// TIA Portal V21 export
// export: Created 2026-11-10T19:11:41.20904Z, ExportSetting WithDefaults, DisplayName Totally Integrated Automation Portal, DisplayVersion V21 Update 3, DisplayName STEP 7 Professional, DisplayVersion V21 Update 3, DisplayName STEP 7 Safety, DisplayVersion V21, DisplayName Tech WebApplication, DisplayVersion V21, DisplayName WinCC Basic/Comfort/Advanced, DisplayVersion V21 Update 3, DisplayName WinCC Unified, DisplayVersion V21 Update 3
DATA_BLOCK "DB_T_CONFIG_SFB"   // DB51
// stored: AutoNumber true, DBAccessibleFromOPCUA true, DBAccessibleFromWebserver true, InstanceOfName T_CONFIG_SFB, OfSystemLibElement T_CONFIG, OfSystemLibVersion 1.0
"T_CONFIG_SFB"
   // VAR_INPUT
   //    Req : Bool;
   //    Interface : HW_INTERFACE;
   //    Conf_Data : Variant;
   // END_VAR
   // VAR_OUTPUT
   //    Done : Bool;
   //    Busy : Bool;
   //    Error : Bool;
   //    Status : DWord;
   //    Err_Loc : DWord;
   // END_VAR
BEGIN
END_DATA_BLOCK
